PROGRAM MAIN
VAR
	comm			: FB_Comm_MQTT_Influx;
	coverControl	: FB_CoverControl(comm := comm);
	focusControl	: FB_FocusControl(comm:=comm);
	haControl		: FB_HourAngleControl(comm:=comm);
	decControl		: FB_DeclinationControl(comm:=comm);
	telescopeControl: FB_TelescopeControl(comm := comm);
	domeControl		: FB_DomeControl(comm := comm);
	pendantControl 	: FB_PendantControl(comm:=comm);
	safetyHandling	: FB_SafetyHandling(comm:=comm);
	rtrigStartUpDone: R_TRIG;
	//search			: FB_RefMarkerSearch(); // use for searching for the Heideinhain encoder reference markers

	
END_VAR
VAR CONSTANT
	telescopeConfig		: ST_TelescopeConfig := (longitude := 9.9452433, latitude := 51.5592378, altitude := 100.0, 
													houranglePark := 0.0, declinationPark := 52.0, focusPark:= 16.3,
													hourangleHome := 0.0, declinationHome := 52.0, focusHome:= 16.3,
													name := 'Emmy Noether', diameter := 0.5, cabinet := 'Beckhoff', manufacturer := '???',
													mountOptions := 'HA-DEC', mount := 'HA_DEC');
END_VAR

//search(Enable:=TRUE); // use for reference marker search

domeControl(ipTelescope	:= telescopeControl);

pendantControl(
	ipTelescope	:= telescopeControl,
	ipFocus		:= focusControl);

coverControl(
	Delta := T#5S,
	TimeToCycle := T#15S,
	bEmergency := safetyHandling.estop);	// previous cycle's value, see bEstopTriggered below (#15)
	
focusControl(
	fVelocity:=1);
	
haControl();
decControl();
telescopeControl(
	fbHourAngle		:= haControl,
	fbDeclination	:= decControl,
	fbFocus			:= focusControl,
	fbDome			:= domeControl,
	fbCovers		:= coverControl,
	telescopeConfig	:= telescopeConfig,
	// was never wired, so STATUS.GLOBAL never reported the E-stop (BROTLib#10). safetyHandling runs below, so
	// this is the previous cycle's value; the drives are cut by the safety circuit regardless.
	bEstopTriggered	:= safetyHandling.estop,
	bSafetyAckPending	:= safetyHandling.ackPending,	// previous cycle, like bEstopTriggered (#59)
);

//Safety
// #11: a telescope reset (cabinet key or the reset command, only fires with an error or a pending acknowledge after an E-stop, #59) also gives the safety
// acknowledge, so the drives leave STO without the VISU
IF telescopeControl.bSafetyAckRequest THEN
	telescopeControl.bSafetyAckRequest := FALSE;
	safetyHandling.Acknowledge();
END_IF
safetyHandling();
// #103: one axis reset pass once the safety start-up is done (the start-up only acknowledges the drives)
rtrigStartUpDone(CLK := safetyHandling.bStartUpDone);
IF rtrigStartUpDone.Q THEN
	telescopeControl.bStartupAxisReset := TRUE;
END_IF

// Comm
comm(	
	sHostName			:= '169.254.149.100',
    nHostPort  			:= 1883,
    nKeepAlive  		:= 10,
	sTopicSub  		 	:= '50cm/Telescope/SET',
	sTopicPublish		:= '50cm/Telemetry',
	sTopicLog			:= '50cm/Log',
	Telescope			:= telescopeControl,
	RaDecTelescope		:= telescopeControl,
	Focus				:= focusControl,
	Dome				:= domeControl,
	MirrorCovers		:= coverControl,
);

END_PROGRAM

(* stored: Version 1.1.0.1, ProductVersion 3.1.4024.15
   POU MAIN: Id {d994e49b-b7f8-4497-8346-561ddfb9c2db}, SpecialFunc None *)
